FUNCTION_BLOCK basicCargaGerador (* Carga alimentada pelos geradores: raio na IHM e bloqueio *)
  (* Standard: 61499-2 *)
  (* Version 1.0, 04/11/2026, Hidryco, Hidryco, 1.0: raio do gerador (0 nao conectado, 1 nao liberada, 2 liberada, 3 liberada e funcionando com a planta nos geradores) e bloqueio (conectada, planta nos geradores e nao liberada na Subestacao). *)
  PACKAGE Hidryco.HidrycoLib;
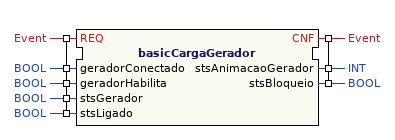
  EVENT_INPUT
    REQ WITH geradorConectado, geradorHabilita, stsGerador, stsLigado; (* Atualizacao *)
  END_EVENT
  EVENT_OUTPUT
    CNF WITH stsAnimacaoGerador, stsBloqueio; (* Raio e bloqueio *)
  END_EVENT
  VAR_INPUT
    geradorConectado : BOOL; (* TRUE = o gerador pode alimentar esta carga *)
    geradorHabilita : BOOL; (* Carga liberada para operar com a planta nos geradores (Subestacao) *)
    stsGerador : BOOL; (* TRUE = planta alimentada pelos geradores *)
    stsLigado : BOOL; (* Carga em funcionamento *)
  END_VAR
  VAR_OUTPUT
    stsAnimacaoGerador : INT; (* 0 nao conectado, 1 nao liberada, 2 liberada, 3 liberada e funcionando nos geradores *)
    stsBloqueio : BOOL; (* Planta nos geradores e carga conectada nao liberada *)
  END_VAR
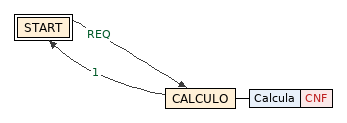
  EC_STATES
    START; (* Estado inicial *)
    CALCULO : Calcula -> CNF; (* Calcula raio e bloqueio *)
  END_STATES
  EC_TRANSITIONS
    START TO CALCULO := REQ;
    CALCULO TO START := 1;
  END_TRANSITIONS
  ALGORITHM Calcula IN ST: (* Raio e bloqueio *)
IF NOT geradorConectado THEN
    stsAnimacaoGerador := 0;
ELSIF NOT geradorHabilita THEN
    stsAnimacaoGerador := 1;
ELSIF stsGerador AND stsLigado THEN
    stsAnimacaoGerador := 3;
ELSE
    stsAnimacaoGerador := 2;
END_IF;
stsBloqueio := geradorConectado AND stsGerador AND NOT geradorHabilita;
  END_ALGORITHM
END_FUNCTION_BLOCK
